VAR_GLOBAL
	Estop1_Y 				AT %I* 	: BOOL ; (* Emergency stop 1 status NC *)
	Estop1_RX 				AT %Q* 	: BOOL ; (* Restart emergency stop NO *)
	
	bLocalEstopFromKUKA 	AT %I* 	: BOOL ;
	bRunStop 				AT %Q*  : BOOL ;
END_VAR

(* stored: Version 1.1.0.1, ProductVersion 3.1.4024.12
   GVL GVL_SAFETY: Id {cad2fc8e-d6ad-422a-a0d5-808b5981c088} *)
